(*
SPDX-FileCopyrightText: © 2026 Oleksandr Tiutyk <trofimich@gmail.com>
SPDX-License-Identifier: MIT
License: https://opensource.org/license/mit
*)

(*!
<summary>Represents an exception raised when a composite activity observes an unexpected child state.</summary>
<description>
Instances are task-scoped diagnostic objects; do not retain references across PLC task cycles.
</description>
*)

INTERFACE IInvalidNestedWorkflowStateException EXTENDS TOF_Core.IGeneralException

(*!
<summary>Formats the invalid nested state diagnostic and raises this exception.</summary>
<description>
Formats bounded diagnostic text without allocating temporary builder storage. Propagation follows the Core
exception lifetime and allocation rules and does not return normally in valid cyclic-task usage.
</description>
<param name="sourceNamespaceName">Namespace of the POU raising the exception.</param>
<param name="sourceClassName">Class name of the composite activity observing the invalid state.</param>
<param name="sourcePOUName">Method or property name where the state was observed.</param>
<param name="sourcePosition">Source position identifier.</param>
<param name="nestedActivityState">Observed child workflow element state that is invalid in the current context.</param>
*)
METHOD Throw
VAR_INPUT
	sourceNamespaceName : STRING;
	sourceClassName : STRING;
	sourcePOUName : STRING;
	sourcePosition : STRING;
	nestedActivityState : WORKFLOW_ELEMENT_STATE;
END_VAR
END_METHOD

END_INTERFACE

(* stored: Version 1.1.0.1
   Itf IInvalidNestedWorkflowStateException: Id {795058f3-1af6-4b6d-a614-ac81afb8e1c0}
   Method Throw: Id {1df65ba3-ad31-4a90-9415-a4bd53aaa136} *)
